Fanuc KAREL source: KD00014.KL

PROGRAM KD00014
%NOLOCKGROUP
VAR
  I: INTEGER
  J: INTEGER
  B: BOOLEAN
  R: REAL
  S: STRING[80]
BEGIN
  RELAX HAND 1
END KD00014
